Yaskawa INFORM job: ENDPOSSEG.JBI

/JOB
//NAME ENDPOSSEG
///FOLDERNAME FOLDER003
//POS
///NPOS 0,0,0,0,0,0
//INST
///DATE 2023/02/17 11:04
///ATTR SC,RW
///GROUP1 RB1
NOP
TIMER T=0.20
SKILLSND "ENDPOSSEG"
ADVINIT
TIMER T=0.20
END
